(* IEC 61131-3 sources: plc-repo-template/src/DUTs, 3 files *)

(* ---- E_DeviceMode.dut.st ---- *)
// Назначение: режимы работы устройства — общие для всех ФБ устройств проекта.
// Автор:      kr0nsch
// Версия:     0.1.0
// Документ:   docs/ARCHITECTURE.md, раздел «Пример в src/»
{attribute 'qualified_only'}
{attribute 'strict'}
TYPE E_DeviceMode :
(
    Auto := 0,          // автоматический: устройством управляет логика ПЛК
    Manual := 1,        // ручной: команды оператора с HMI/SCADA
    Local := 2,         // местный: управление с местного поста, команда ПЛК снимается
    OutOfService := 3   // выведено из работы: выход в безопасном состоянии, команды игнорируются
);
END_TYPE

(* ---- ST_ExampleCmd.dut.st ---- *)
// Назначение: команды HMI/SCADA для примера FB_Example (насос подкачки).
//             Однократные команды (xAck, xReset) сбрасывает ПЛК после выполнения.
// Автор:      kr0nsch
// Версия:     0.1.0
// Документ:   docs/ARCHITECTURE.md, раздел «Пример в src/»
TYPE ST_ExampleCmd :
STRUCT
    // требуемый режим; после холодного старта устройство выведено из работы
    eMode : E_DeviceMode := E_DeviceMode.OutOfService;
    // уставка отключения, % диапазона датчика
    rSetpoint_pct : REAL := GVL_Const.EXAMPLE_SP_DEFAULT_PCT;
    xManualOn : BOOL;       // ручная команда «включить» (режим Manual)
    xAck : BOOL;            // квитирование отказа (однократная команда)
    xReset : BOOL;          // сброс состояния и счётчика (однократная команда)
END_STRUCT
END_TYPE

(* ---- ST_ExampleSts.dut.st ---- *)
// Назначение: состояние примера FB_Example для HMI/SCADA.
// Автор:      kr0nsch
// Версия:     0.1.0
// Документ:   docs/ARCHITECTURE.md, раздел «Пример в src/»
TYPE ST_ExampleSts :
STRUCT
    eMode : E_DeviceMode;           // действующий режим
    xOut : BOOL;                    // выход включён
    xFault : BOOL;                  // отказ измерения зафиксирован, ждёт квитирования
    rSetpointUsed_pct : REAL;       // действующая уставка после ограничения, %
    udiCount : UDINT;               // число включений выхода с последнего сброса
END_STRUCT
END_TYPE
